// TIA Portal V19 export
TYPE "PidL.Permission"
   STRUCT
      AutModOpEn : Bool;
      ManModOpEn : Bool;
      LocModOpEn : Bool;
      OosModOpEn : Bool;
      ResetOpEn : Bool;
      ExtModOpEn : Bool;
      IntModOpEn : Bool;
      Alarms { S7_SetPoint := 'True'} : "AnaMon.Permission";
   END_STRUCT;
END_TYPE
